INTERFACE I_Station EXTENDS __SYSTEM.IQueryInterface

METHOD HasMover : BOOL
VAR_INPUT
END_VAR
END_METHOD

METHOD IsClear : BOOL
VAR_INPUT
END_VAR
END_METHOD

METHOD isComplete : BOOL
VAR_INPUT
END_VAR
END_METHOD

METHOD IsOperating : BOOL
VAR_INPUT
END_VAR
END_METHOD

METHOD IsReady : BOOL
VAR_INPUT
END_VAR
END_METHOD

METHOD MyMover : HRESULT
VAR_INPUT
	mover : I_XtsMover;
END_VAR
END_METHOD

PROPERTY Position : MC_LREAL
GET
END_GET
END_PROPERTY

END_INTERFACE

(* stored: Version 1.1.0.1
   Itf I_Station: Id {d8773b48-8571-4ecd-8cbd-ba8942597bd4}
   Method HasMover: Id {5b7781a3-78e4-4116-9d74-37fb48cc3c12}
   Method IsClear: Id {3b338444-496f-4b57-aaf3-4efffa633361}
   Method isComplete: Id {60ede7f6-c745-40a4-bf92-f3a03a7a1452}
   Method IsOperating: Id {e04f481b-64f7-4cd5-aead-d2162ca18486}
   Method IsReady: Id {1429945e-e662-41b3-82dc-271da72170fa}
   Method MyMover: Id {e0d36098-8d65-476a-990c-e6fc9c4a3a40}
   Property Position: Id {382268c5-e001-4500-92a7-4729d1276a58}
   Get Get: Id {419af852-7c98-4df9-a521-739afc5b0cdd} *)
